DATA_BLOCK "S11RecoveryGraph"
{ S7_Optimized_Access := 'TRUE' }
VERSION : 0.1
NON_RETAIN
"FB_S11RecoveryGraph"
BEGIN
END_DATA_BLOCK
